(* Schneider Machine Expert - Basic project ECE4311_PLC, file version 3.0.0.0 *)
(* CompanyInformations: Name=CPP *)
(* ProjectInformations: Name=ControlShield, Description=ECE4311 – Network Forensics: Development of a PLC Guardian HMI for the M221 PLC on an HMIS5T panel, focusing on cybersecurity and network forensics for industrial control systems. *)

HARDWARE
  Cpu 0: TM221CE24T
  EthernetConfiguration: NetworkName=M221, IpAllocationMode=FixedAddress, IpAddress=192.168.8.11, SubnetMask=255.255.255.0
  SerialLineConfiguration: Baud=Baud19200, Parity=ParityEven, DataBits=DataBits8, StopBits=StopBits1, PhysicalMedium=PhysicalMediumRs485, TransmissionMode=TransmissionModeModbusRtu, SlaveId=1, Addressing=SlaveAddressing
  MastTask: UsePeriodScanMode=false, PeriodScan=100
  FastTask: Period=255
  CpuBehavior: StartingMode=StartAsPreviousState, AutoSaveRamOnEeprom=true, WatchdogPeriod=250

SYMBOLS  (address, symbol, comment, settings)
  %M0       T1
  %M1       T2
  %M2       STARTBUTTON
  %M3       STOP
  %M4       MAINT_BYPASS
  %M5       RESET
  %M6       DIGI_OVERLOAD
  %MW0      TANK_VALUE
  %TM0      TICK  [Preset=100, Base=OneMilliSeconds]
  %TM1      TOCK  [Type=TOF, Preset=100, Base=OneMilliSeconds]
  %C0       TANK_N  [Preset=80]
  %Q0.0     OUTPUT_1
  %Q0.1     OUTPUT_2
  %Q0.2     TANK_OVERLOAD

POU Main
  (* SectionNumber=1 *)

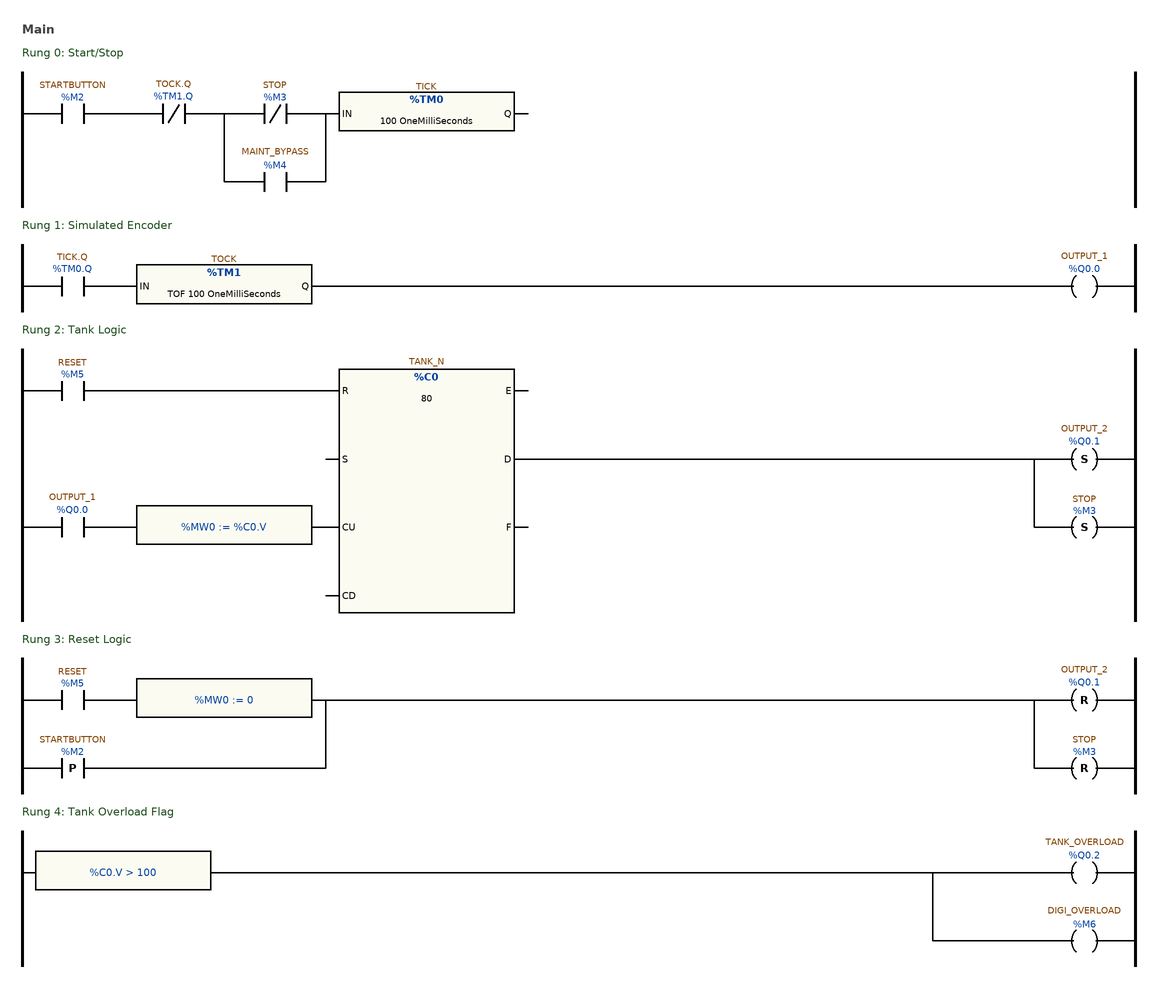

// Rung 0: Start/Stop
  BLK %TM0                (* TICK *)
  LD %M2                  (* STARTBUTTON *)
  ANDN %TM1.Q             (* TOCK *)
  AND(N %M3               (* STOP *)
  OR %M4                  (* MAINT_BYPASS *)
  )
  IN
  END_BLK
  // as ST:
  //   TICK(IN := STARTBUTTON AND NOT TOCK.Q AND (NOT STOP OR MAINT_BYPASS));

// Rung 1: Simulated Encoder
  BLK %TM1                (* TOCK *)
  LD %TM0.Q               (* TICK *)
  IN
  OUT_BLK
  LD Q
  ST %Q0.0                (* OUTPUT_1 *)
  END_BLK
  // as ST:
  //   TOCK(IN := TICK.Q);
  //   OUTPUT_1 := TOCK.Q;

// Rung 2: Tank Logic
  BLK %C0                 (* TANK_N *)
  LD %M5                  (* RESET *)
  R
  LD %Q0.0                (* OUTPUT_1 *)
  OPER [ %MW0 := %C0.V ]  (* TANK_VALUE, TANK_N *)
  CU
  OUT_BLK
  LD D
  S %Q0.1                 (* OUTPUT_2 *)
  S %M3                   (* STOP *)
  END_BLK
  // as ST:
  //   IF OUTPUT_1 THEN TANK_VALUE := TANK_N.V; END_IF;
  //   TANK_N(R := RESET, CU := OUTPUT_1);
  //   IF TANK_N.D THEN OUTPUT_2 := TRUE; END_IF;
  //   IF TANK_N.D THEN STOP := TRUE; END_IF;

// Rung 3: Reset Logic
  LD %M5                  (* RESET *)
  OPER [ %MW0 := 0 ]      (* TANK_VALUE *)
  ORR %M2                 (* STARTBUTTON *)
  R %Q0.1                 (* OUTPUT_2 *)
  R %M3                   (* STOP *)
  // as ST:
  //   IF RESET THEN TANK_VALUE := 0; END_IF;
  //   IF RESET OR RISING(STARTBUTTON) THEN OUTPUT_2 := FALSE; END_IF;
  //   IF RESET OR RISING(STARTBUTTON) THEN STOP := FALSE; END_IF;

// Rung 4: Tank Overload Flag
  LD [ %C0.V > 100 ]      (* TANK_N *)
  ST %Q0.2                (* TANK_OVERLOAD *)
  ST %M6                  (* DIGI_OVERLOAD *)
  // as ST:
  //   TANK_OVERLOAD := TANK_N.V > 100;
  //   DIGI_OVERLOAD := TANK_N.V > 100;
